Staubli VAL3: modifyFrame.pgx

program modifyFrame(num x_nIndex)
  local bool l_bExit
  local num l_i
  local string l_sNmb
begin
  do
    if util:sPage!="frameSetting"
      util:sPage="frameSetting"

      nFrame[0]=savedata:fFrameItem[x_nIndex].fFrame.trsf.x
      nFrame[1]=savedata:fFrameItem[x_nIndex].fFrame.trsf.y
      nFrame[2]=savedata:fFrameItem[x_nIndex].fFrame.trsf.z
      nFrame[3]=savedata:fFrameItem[x_nIndex].fFrame.trsf.rx
      nFrame[4]=savedata:fFrameItem[x_nIndex].fFrame.trsf.ry
      nFrame[5]=savedata:fFrameItem[x_nIndex].fFrame.trsf.rz
      for l_i = 0 to 5
        l_sNmb="nmb"+toString("",l_i+1)
        userPageBind("frameSetting",l_sNmb,"value",nFrame[l_i],1,"rw")
      endFor
      userPageBindClick("frameSetting","btn1",bModifyFrame,true)
      userPageBindClick("frameSetting","btn2",bCancelFrame,true)
      userPage(util:sPage)
      delay(0.5)
    endIf

    if bModifyFrame
      bModifyFrame=false
      savedata:fFrameItem[x_nIndex].fFrame.trsf.x=nFrame[0]
      savedata:fFrameItem[x_nIndex].fFrame.trsf.y=nFrame[1]
      savedata:fFrameItem[x_nIndex].fFrame.trsf.z=nFrame[2]
      savedata:fFrameItem[x_nIndex].fFrame.trsf.rx=nFrame[3]
      savedata:fFrameItem[x_nIndex].fFrame.trsf.ry=nFrame[4]
      savedata:fFrameItem[x_nIndex].fFrame.trsf.rz=nFrame[5]
      savedata:libSave()
      delay(0.1)
       l_bExit=true
    elseIf bCancelFrame
      bCancelFrame=false
      l_bExit=true
    endIf
    delay(0)
  until l_bExit==true
end
